Staubli VAL3: insertJoint.pgx

public program insertJoint(string x_sKey, num x_nIndex, bool& x_bToSave)
  local num l_j
  local num l_i
begin
  // insert(trajTemp:tTrajItem[x_sKey].pPointItem[x_nIndex+1])
  append(trajTemp:tTrajItem[x_sKey].pPointItem)

  for l_i = (size(trajTemp:tTrajItem[x_sKey].pPointItem)-1) to(x_nIndex+1) step -1
    //logMsg(toString("",l_i))
    call copyPoint3(x_sKey,l_i,l_i-1)
  endFor
  trajTemp:tTrajItem[x_sKey].pPointItem[x_nIndex+1].pPointRx=trajTemp:tTrajItem[x_sKey].pPointItem[x_nIndex].pPointRx
  trajTemp:tTrajItem[x_sKey].pPointItem[x_nIndex+1].jJointRx=trajTemp:tTrajItem[x_sKey].pPointItem[x_nIndex].jJointRx
  trajTemp:tTrajItem[x_sKey].pPointItem[x_nIndex+1].pParaItem.mMdesc=trajTemp:tTrajItem[x_sKey].pPointItem[x_nIndex].pParaItem.mMdesc
  trajTemp:tTrajItem[x_sKey].pPointItem[x_nIndex+1].pParaItem.nMoveType=0
  trajTemp:tTrajItem[x_sKey].pPointItem[x_nIndex+1].pParaItem.nDelay=trajTemp:tTrajItem[x_sKey].pPointItem[x_nIndex].pParaItem.nDelay
  trajTemp:tTrajItem[x_sKey].pPointItem[x_nIndex+1].pParaItem.nSigValue=trajTemp:tTrajItem[x_sKey].pPointItem[x_nIndex].pParaItem.nSigValue
  trajTemp:tTrajItem[x_sKey].pPointItem[x_nIndex+1].pParaItem.nActionIndex=trajTemp:tTrajItem[x_sKey].pPointItem[x_nIndex].pParaItem.nActionIndex
  trajTemp:tTrajItem[x_sKey].pPointItem[x_nIndex+1].pParaItem.nPercentage=trajTemp:tTrajItem[x_sKey].pPointItem[x_nIndex].pParaItem.nPercentage
  for l_j = 0 to 2
    trajTemp:tTrajItem[x_sKey].pPointItem[x_nIndex+1].pParaItem.iIfItem.nSigType[l_j]=trajTemp:tTrajItem[x_sKey].pPointItem[x_nIndex].pParaItem.iIfItem.nSigType[l_j]
    trajTemp:tTrajItem[x_sKey].pPointItem[x_nIndex+1].pParaItem.iIfItem.nSigIndex[l_j]=trajTemp:tTrajItem[x_sKey].pPointItem[x_nIndex].pParaItem.iIfItem.nSigIndex[l_j]
    trajTemp:tTrajItem[x_sKey].pPointItem[x_nIndex+1].pParaItem.iIfItem.nValue[l_j]=trajTemp:tTrajItem[x_sKey].pPointItem[x_nIndex].pParaItem.iIfItem.nValue[l_j]
  endFor
  //trajTemp:libSave()
  x_bToSave=true
end
